Staubli VAL3: waitAnaInput.pgx

public program waitAnaInput(aio x_aIn, num x_nValue, bool& x_bError)
  local string l_sDesc
  local string l_sPath
begin
  if ioStatus(x_aIn,l_sDesc,l_sPath)>=0
    x_bError=false
    wait(aioGet(x_aIn)==x_nValue)
  else
    x_bError=true
    logMsg("通信终端，等待通信恢复")
    wait(aioGet(x_aIn)==x_nValue)
    logMsg("通信已恢复")
    //    logMsg("Signal "+l_sPath+" error."+"Description:"+l_sDesc)
  endIf
end
